(* IEC 61131-3 sources: model-first-plc-agent-ai/results/T2-W-02, 2 files *)

(* ---- a1_code.st ---- *)
FUNCTION_BLOCK FillingRuntime
VAR_INPUT
    start : BOOL;
    stop : BOOL;
    LSH : BOOL;
    LSHH : BOOL;
    TimerDuration : TIME;
END_VAR
VAR_OUTPUT
    fill_valve : BOOL;
    discharge_valve : BOOL;
END_VAR
VAR
    ActiveState : INT := 0;
    FillingTimer : TON;
    timer_done : BOOL := FALSE;
END_VAR

CASE ActiveState OF
    0:
        timer_done := FALSE;

        IF start AND NOT stop AND NOT LSHH THEN
            ActiveState := 1;
        END_IF;

        (* Start timing in the scan that activates x1. *)
        FillingTimer(
            IN := (ActiveState = 1),
            PT := TimerDuration
        );

    1:
        FillingTimer(IN := TRUE, PT := TimerDuration);
        timer_done := FillingTimer.Q;

        IF stop OR LSHH OR timer_done THEN
            ActiveState := 0;
            FillingTimer(IN := FALSE, PT := TimerDuration);
            timer_done := FALSE;
        END_IF;

ELSE
    ActiveState := 0;
    FillingTimer(IN := FALSE, PT := TimerDuration);
    timer_done := FALSE;
END_CASE;

fill_valve := (ActiveState = 1);
discharge_valve := FALSE;

END_FUNCTION_BLOCK

PROGRAM Main
VAR
    StartCommand AT %IX100.0 : BOOL;
    StopCommand AT %IX100.1 : BOOL;
    LSH AT %IX100.2 : BOOL;
    LSHH AT %IX100.3 : BOOL;

    FillValve AT %QX100.0 : BOOL;
    DischargeValve AT %QX100.1 : BOOL;
END_VAR
VAR
    (* Configurable filling interval; example initial setting. *)
    TimerDuration : TIME := T#10s;
    StartEdge : R_TRIG;
    Controller : FillingRuntime;
END_VAR

StartEdge(CLK := StartCommand);

Controller(
    start := StartEdge.Q,
    stop := StopCommand,
    LSH := LSH,
    LSHH := LSHH,
    TimerDuration := TimerDuration
);

FillValve := Controller.fill_valve;
DischargeValve := Controller.discharge_valve;

END_PROGRAM

(* ---- a2_code.st ---- *)
FUNCTION_BLOCK FB_TimedTank
VAR_INPUT
    StartCommand : BOOL;
    StopCommand : BOOL;
    LSH : BOOL;
    LSHH : BOOL;
    TimerDuration : TIME;
END_VAR
VAR_OUTPUT
    fill_valve : BOOL;
    discharge_valve : BOOL;
END_VAR
VAR
    StartEdge : R_TRIG;
    FillingTimer : TON;
    start : BOOL;
    stop : BOOL;
    timer_done : BOOL;
    x1 : BOOL := FALSE;
END_VAR

(* Detect each press, including presses during stop or filling. *)
StartEdge(CLK := StartCommand);
start := StartEdge.Q;
stop := StopCommand;

(* Stop and high-high detection take priority over starting. *)
IF stop OR LSHH THEN
    x1 := FALSE;
ELSIF NOT x1 AND start THEN
    x1 := TRUE;
END_IF;

(* Timing begins in the same scan as entry into the filling step. *)
FillingTimer(IN := x1, PT := TimerDuration);
timer_done := FillingTimer.Q;

IF x1 AND timer_done THEN
    x1 := FALSE;

    (* Reset the owned timer immediately on leaving its step. *)
    FillingTimer(IN := FALSE, PT := TimerDuration);
    timer_done := FillingTimer.Q;
END_IF;

fill_valve := x1;
discharge_valve := FALSE;

END_FUNCTION_BLOCK

PROGRAM Main
VAR
    StartCommand AT %IX100.0 : BOOL;
    StopCommand AT %IX100.1 : BOOL;
    LSH AT %IX100.2 : BOOL;
    LSHH AT %IX100.3 : BOOL;
    FillValve AT %QX100.0 : BOOL;
    DischargeValve AT %QX100.1 : BOOL;
END_VAR
VAR
    TankController : FB_TimedTank;
    (* Configurable preset; adjust to the required filling duration. *)
    TimerDuration : TIME := T#10s;
END_VAR

TankController(
    StartCommand := StartCommand,
    StopCommand := StopCommand,
    LSH := LSH,
    LSHH := LSHH,
    TimerDuration := TimerDuration
);

FillValve := TankController.fill_valve;
DischargeValve := TankController.discharge_valve;

END_PROGRAM
